TYPE ST_UDPFrameEntry :
STRUCT
	stRemoteAddr 	: ST_SockAddr;	(* Remote address. String containing an (Ipv4) Internet Protocol dotted address and port number. *)
	sMessage		: UDP_DATA;	(* UDP packet data *)
END_STRUCT
END_TYPE

(* stored: Version 1.1.0.1
   DUT ST_UDPFrameEntry: Id {02fc53d0-13a1-413a-bb04-7ebaa8d43742} *)
